Staubli VAL3: autoReturn.dtx

mdesc mNomSpeed
public num nRecIndex
num nMoveIdRec[200]
trsf trToolRec[200]
jointRx jPointRec[200 2]
num nMoveTypeRec[200]
mdesc mReturn = {accel=5, vel=10, decel=5, leave=1, reach=1}
bool bFirstUpdate
mdesc mSpeedRec[200]
jointRx jRefPoint
num nRefDeviate
bool bPushToStack
bool bExact[200]
num nCurrentMoveID
public bool bInterrupt
num nIndex
bool bHaveGetMoveID
